(*~
		<docu>
			<summary>
				Provides mechanism for delivering static messages to the supervising applications (SCADA/HMI).	
				<remarks>			
					<note type="important">
						Each messenger has a single placeholder for the message; it stores the most important message from the last context cycle. 
						If there are more messages in a single cycle for the same messenger then less important messages are discarded and replaced by 
						the message with the category of higher severity.							
					</note>
					<note type="important">
						Messenger can send the data to context logger. There is a maximum limit of 10 different messages per messenger in 2 consecutive context cycles.
						The messages that exceed this limit won't be logged when `OnEventRisen` logging is set. 
					    Take this behaviour into account when designing your system.				
					</note>					
				</remarks>			 
			</summary>			
		
		</docu>
~*)
FUNCTION_BLOCK PUBLIC TcoMessenger IMPLEMENTS ITcoMessenger, ITcoMessageProperties, ITcoMessageTextBuilder, ITcoMessageCategorize
VAR			
	(*~
		<docu>
			<summary>
				Most important message of this instance of messenger; stores the most important message from the last context cycle. 
				If there are more messages in a single cycle for the same
				messenger then less important messages are discarded and replaced by the message with the category of higher severity.			 
			</summary>			
		</docu>
	~*)
	_mime : TcoMessage;
	_Parent : ITcoObject;
	{attribute clr [ReadOnly()]}
	_contextIdentity : ULINT;	
	{attribute 'hide'}
	_mds : ARRAY[0..MDS_MAX_INDEX] OF TcoMessageDigest;	
	{attribute 'hide'}
	_condition : eMessageCondition;
	{attribute 'hide'}
	_pinnable : BOOL;		
END_VAR

VAR
	{attribute 'hide'}
	tmpMessageText : STRING(TcoMessengerEnv.MAX_MESSAGE_TEXT_LENGHT);
	{attribute 'hide'}
	refStringBuilder : REFERENCE TO StringBuilder;	
END_VAR

VAR CONSTANT
	MDS_MAX_INDEX : INT := 10;
END_VAR

VAR_STAT
	{attribute 'hide'}
	_conflictingStringBuilder : StringBuilder;
END_VAR

(*~
	<docu>
		<summary>			
			Appends string to the message text. 
		</summary>
		<remarks>
			<note type="warning">
				The size of the resulting string should not be more than '160' characters. The characters exceeding this size will be truncated.
			</note>
		</remarks>
	</docu>	
~*)
{attribute 'hide'}
{attribute 'obsolete' := 'This method must be accessed ITcoMessageTextBuilder interface'} 
METHOD Append : ITcoMessageTextBuilder
VAR_INPUT
	Text : STRING(TcoMessengerEnv.MAX_MESSAGE_TEXT_LENGHT);
END_VAR
THIS^.StringBuilder.Append(Text);
Append := THIS^;
END_METHOD

(*~
	<docu>
		<summary>			
			Appends any value to the message text. 
		</summary>
		<remarks>
			<note type="warning">
				The size of the resulting string should not be more than '160' characters. The characters exceeding this size will be truncated.
			</note>
		</remarks>
	</docu>	
~*)
METHOD AppendAny : ITcoMessageTextBuilder
VAR_INPUT
	Data : ANY;
END_VAR
THIS^.StringBuilder.AppendAny(Data);
AppendAny := THIS^;
END_METHOD

(*~
	<docu>
		<summary>			
			Gets categorization methods for fluent message builder.
		</summary>		
	</docu>	
~*)
{attribute 'hide'}
{attribute 'obsolete' := 'This method must be accessed ITcoMessageTextBuilder interface'} 
METHOD As : ITcoMessageCategorize
As := THIS^;
END_METHOD

(*~
		<docu>
			<summary>
				Categotizes and creates the message as  'debug'.								 
			</summary>		
		</docu>
~*)
{attribute 'hide'}
{attribute 'obsolete' := 'This method must be accessed ITcoMessageCategorize interface'} 
METHOD PUBLIC AsDebug : ITcoMessageProperties
AsDebug := Post(THIS^.StringBuilder.ToString(), eMessageCategory.Debug);
END_METHOD

(*~
		<docu>
			<summary>
				Categotizes and creates the message as  'error'.								 
			</summary>		
		</docu>
~*)

{attribute 'hide'}
{attribute 'obsolete' := 'This method must be accessed ITcoMessageCategorize interface'} 
METHOD PUBLIC AsError : ITcoMessageProperties
AsError := Post(THIS^.StringBuilder.ToString(), eMessageCategory.Error);
END_METHOD

(*~
		<docu>
			<summary>
				Categotizes and creates the message as  'fatal'.								 
			</summary>		
		</docu>
~*)

{attribute 'hide'}
{attribute 'obsolete' := 'This method must be accessed ITcoMessageCategorize interface'} 
METHOD PUBLIC AsFatal : ITcoMessageProperties
AsFatal := Post(THIS^.StringBuilder.ToString(), eMessageCategory.Fatal);
END_METHOD

(*~
		<docu>
			<summary>
				Categotizes and creates the message as  'information'.								 
			</summary>		
		</docu>
~*)

{attribute 'hide'}
{attribute 'obsolete' := 'This method must be accessed ITcoMessageCategorize interface'} 
METHOD PUBLIC AsInfo : ITcoMessageProperties
AsInfo := Post(THIS^.StringBuilder.ToString(), eMessageCategory.Info);
END_METHOD

(*~
		<docu>
			<summary>
				Categotizes and creates the message as  'trace'.								 
			</summary>		
		</docu>
~*)

{attribute 'hide'}
{attribute 'obsolete' := 'This method must be accessed ITcoMessageCategorize interface'} 
METHOD PUBLIC AsTrace : ITcoMessageProperties
AsTrace := Post(THIS^.StringBuilder.ToString(), eMessageCategory.Trace);
END_METHOD

(*~
		<docu>
			<summary>
				Categotizes and creates the message as 'warning'.								 
			</summary>		
		</docu>
~*)

{attribute 'hide'}
{attribute 'obsolete' := 'This method must be accessed ITcoMessageCategorize interface'} 
METHOD PUBLIC AsWarning : ITcoMessageProperties
AsWarning := Post(THIS^.StringBuilder.ToString(), eMessageCategory.Warning);
END_METHOD

(*~
	<docu>
		<summary>			
			Initiates new message text building for this messenger in fluent-like fashion.
		</summary>		
	</docu>	
~*)
METHOD Build : ITcoMessageTextBuilder
THIS^.StringBuilder.Clear();
Build := THIS^;
END_METHOD

(*~
		<docu>
			<summary>
				Adds message of 'catastrophic' category to the message queue.
				Use this category when there is a situation when the device cannot continue operations due to irrecoverable failure.				 
			</summary>		
		</docu>
~*)
METHOD PUBLIC Catastrophic : ITcoMessageProperties
VAR_INPUT
	(*~
		<docu>
			<summary>
				Arbitrary message string.			 
			</summary>			
		</docu>
	~*)
	Message : STRING(TcoMessengerEnv.MAX_MESSAGE_TEXT_LENGHT);
END_VAR
Catastrophic := THIS^.Post(Message, eMessageCategory.Catastrophic);
END_METHOD

(*~
		<docu>
			<summary>
				Clears the message content.
				<remarks>			
					<note type="important">
						This method is exposed for Rpc calls, for testing purposes. Rpc calls of this method must not be used in production code
					</note>
				</remarks>								 
			</summary>		
		</docu>
~*)
{attribute 'TcRpcEnable'}
METHOD Clear
_mime.TimeStamp :=  DT#1970-01-01-00:00;
_mime.Text := '';
_mime.Identity := 0;
_mime.Category := eMessageCategory.All;
_mime.Cycle := 0;	
_mime.PerCycleCount := 0;
_mime.Pinned := FALSE;
END_METHOD

METHOD PROTECTED Compose : TcoMessage
VAR_INPUT
	Text : STRING(TcoMessengerEnv.MAX_MESSAGE_TEXT_LENGHT);
	Category : eMessageCategory;
END_VAR
IF(_Parent <> 0 AND_THEN _Parent.Context <> 0 AND_THEN _Parent.Context.RealTimeClock <> 0) THEN
	Compose.TimeStamp :=  _Parent.Context.RealTimeClock.NowLocal();	
	Compose.Text := Text;
	Compose.Identity := _Parent.Identity;
	Compose.Category := Category;
	Compose.Cycle := _Parent.Context.StartCycleCount;
	Compose.MessageDigest := Digest(Text, THIS^._Parent.Context.Environment.Messaging.MessageDigestMethod);
END_IF;
END_METHOD

(*~
		<docu>
			<summary>
				Adds message of 'critical' category to the message queue.
				Use this category when a critical error occured, that is not recoverable by the means of software (reset/restore) and a detailed inspection is required.				 
			</summary>		
		</docu>
~*)
METHOD PUBLIC Critical : ITcoMessageProperties
VAR_INPUT
	(*~
		<docu>
			<summary>
				Arbitrary message string.			 
			</summary>			
		</docu>
	~*)
	Message : STRING(TcoMessengerEnv.MAX_MESSAGE_TEXT_LENGHT);
END_VAR
Critical := THIS^.Post(Message, eMessageCategory.Critical);
END_METHOD

(*~
		<docu>
			<summary>
				Adds message of 'debug' category to the message queue.	
			    Use when you need to report debug information for you as programmer. 			 
			</summary>		
		</docu>
~*)
METHOD PUBLIC Debug : ITcoMessageProperties
VAR_INPUT
	(*~
		<docu>
			<summary>
				Arbitrary message string.			 
			</summary>			
		</docu>
	~*)
	Message : STRING(TcoMessengerEnv.MAX_MESSAGE_TEXT_LENGHT);
END_VAR
Debug := THIS^.Post(Message, eMessageCategory.Debug);
END_METHOD

METHOD Digest : DWORD
VAR_INPUT
	Text : Tc2_System.T_MaxString;
	inDigestType : eMessageDigestMethod;
END_VAR
CASE inDigestType OF
	eMessageDigestMethod.CRC8 :
		Digest := TcoCRC_8(Text);
	eMessageDigestMethod.CRC16 :
		Digest := TcoCRC_16(Text);
	eMessageDigestMethod.CRC32 :
		Digest := TcoCRC_32(Text);
	ELSE
		Digest := 0;
END_CASE
END_METHOD

(*~
		<docu>
			<summary>
				Adds message of 'error' category to the message queue.
				Use this categoty when there is a failure that cannot be immediately recovered and an intervention is needed. This is typically a situation when a device fails
				to deliver expected result. 
				Do not use this category to report information about failed process like measurement or detection.				 
			</summary>						
		</docu>
~*)
METHOD PUBLIC Error : ITcoMessageProperties
VAR_INPUT
	(*~
		<docu>
			<summary>
				Arbitrary message string.			 
			</summary>			
		</docu>
	~*)
	Message : STRING(TcoMessengerEnv.MAX_MESSAGE_TEXT_LENGHT);
END_VAR
Error := THIS^.Post(Message, eMessageCategory.Error);
END_METHOD

{attribute 'hide'}
METHOD FB_init : BOOL
VAR_INPUT
	bInitRetains : BOOL; // if TRUE, the retain variables are initialized (warm start / cold start)
	bInCopyCode : BOOL;  // if TRUE, the instance afterwards gets moved into the copy code (online change)
	ParentObject : ITcoObject;
END_VAR
_Parent := ParentObject;
_contextIdentity := ParentObject.Identity;
END_METHOD

(*~
		<docu>
			<summary>
				Adds message of 'information' category to the message queue.	
				Use when you want to deliver information to the user, that has only informative character and does not adversely affect a process.			 
			</summary>			
		</docu>
~*)
METHOD PUBLIC Info  : ITcoMessageProperties
VAR_INPUT
	(*~
		<docu>
			<summary>
				Arbitrary message string.			 
			</summary>			
		</docu>
	~*)
	Message : STRING(TcoMessengerEnv.MAX_MESSAGE_TEXT_LENGHT);
END_VAR
Info := THIS^.Post(Message, eMessageCategory.Info);
END_METHOD

METHOD PRIVATE LogMessage 
VAR_IN_OUT
	inMessage : TcoMessage;
END_VAR
VAR
	_index : INT;
	_freeIndex : INT;	
END_VAR
CASE _Parent.Context.Environment.Messaging.MessengerLoggingMethod OF
	eMessengerLogMethod.OnEventRisen :
        IF(_Parent.Context.Environment.Messaging.MessageDigestMethod = eMessageDigestMethod.NONE) THEN
			inMessage.MessageDigest := Digest(inMessage.Text, eMessageDigestMethod.CRC32);
		END_IF
	
		_freeIndex := 0;
		    
		FOR _index := 0 TO MDS_MAX_INDEX DO
			IF(_mds[_index].Cycle = inMessage.Cycle - 1 OR _mds[_index].Cycle = inMessage.Cycle) 
			AND_THEN (_mds[_index].Digest = inMessage.MessageDigest)
			AND_THEN (_mds[_index].Category = inMessage.Category) THEN			
			    _mds[_index].Cycle := inMessage.Cycle;				
				RETURN;											
			END_IF	
			IF((_mds[_index].Cycle <> inMessage.Cycle - 1) 
			   AND (_mds[_index].Cycle <> inMessage.Cycle)) THEN
				_freeIndex := _index;
			END_IF
		END_FOR
		
		IF(_freeIndex <= THIS^.MDS_MAX_INDEX) THEN
			_mds[_freeIndex].Digest := inMessage.MessageDigest;
			_mds[_freeIndex].Cycle := inMessage.Cycle;
			_mds[_freeIndex].Category := inMessage.Category;
			_Parent.Context.Logger.PushMessage(inMessage);		
		END_IF;
	eMessengerLogMethod.Continuous:
	    _Parent.Context.Logger.PushMessage(inMessage);
END_CASE
END_METHOD

(*~
		<docu>
			<summary>
				Adds message of 'notification' category to the message queue.
				Use this category when you want to report a notification that may be of interest to the user, but does not adveresly affect a process.			 
			</summary>				
		</docu>
~*)
METHOD Notify : ITcoMessageProperties
VAR_INPUT
	(*~
		<docu>
			<summary>
				Arbitrary message string.			 
			</summary>			
		</docu>
	~*)
	Message : STRING(TcoMessengerEnv.MAX_MESSAGE_TEXT_LENGHT);
END_VAR
Notify := THIS^.Post(Message, eMessageCategory.Notification);
END_METHOD

METHOD OnCondition : ITcoMessages
VAR_INPUT
	inCondition : BOOL;
END_VAR
IF (inCondition) THEN
	_condition := eMessageCondition.Active;
ELSE
	_condition := eMessageCondition.Inactive;
END_IF

OnCondition := THIS^;
END_METHOD

(*~
	<docu>
		<summary>
			Pins this message that no other message will override it. 
			The messenger won't accept new messages until acknowledged in diagnostics view by user, unipenned by `Unpin()` methods or cleared by `Clear()` method
			of this messenger.						
		</summary>
		<note type="important">
			Pinned messages do no accept incomming messages on the same messenger. The incomming messages will be though the context logger when active.
		</note>
	</docu>
~*)
//~
{attribute 'hide'}
{attribute 'obsolete' := 'This method must be called exclusively over ITcoMessageProperties interface'}
//~ 
METHOD Pin : ITcoMessageProperties
IF(_Parent <> 0 AND_THEN _Parent.Context <> 0) THEN
	IF(_pinnable AND_THEN _mime.Cycle = _Parent.Context.StartCycleCount)THEN
		_mime.Pinned := TRUE;
	END_IF;
END_IF;

Pin := THIS^;
END_METHOD

(*~
	<docu>
		<summary>
			Gets `true` when this messanger is pinned (awaiting acknowledgement in diagnostics view).
		</summary>
	</docu>
~*)
PROPERTY Pinned : BOOL
GET
Pinned := _mime.Pinned AND_THEN tmpMessageText = _mime.Text;
END_GET
END_PROPERTY

(*~
		<docu>
			<summary>
				Creates message of given category for this messenger.				 
			</summary>				
		</docu>
~*)
METHOD PUBLIC Post : ITcoMessageProperties
VAR_INPUT
	(*~
		<docu>
			<summary>
				Arbitrary message string.			 
			</summary>			
		</docu>
	~*)
	Message : STRING(TcoMessengerEnv.MAX_MESSAGE_TEXT_LENGHT);
	(*~
		<docu>
			<summary>
				Message category.			 
			</summary>			
		</docu>
	~*)
	Category : eMessageCategory;	
END_VAR

VAR
	_wouldBeMime : TcoMessage;
END_VAR
Post := THIS^;

tmpMessageText := Message;

_pinnable := FALSE;

IF(_condition = eMessageCondition.Inactive) THEN
	_condition := eMessageCondition.Unconditional;	
	RETURN;
END_IF

_condition := eMessageCondition.Unconditional;


IF(_Parent <> 0 AND_THEN _Parent.Context <> 0 AND_THEN _Parent.Context.Environment <> 0 AND_THEN _Parent.Context.Environment.Messaging <> 0) THEN
	IF(Category < THIS^._Parent.Context.Environment.Messaging.MinLevel
	  OR _Parent.Context.Environment.Messaging.IsSuspended) THEN
		RETURN;
	END_IF; 	
		
	IF (NOT _mime.Pinned) THEN 
		_mime.PerCycleCount := _mime.PerCycleCount + 1;
		_wouldBeMime := Compose(Message, Category);		
		_wouldBeMime.PerCycleCount := _mime.PerCycleCount;		
	ELSIF(_mime.Pinned 
	AND_THEN (_mime.Text <>  Message OR _mime.Category <> Category))
	THEN		
		IF(	_mime.PerCycleCount < 255) THEN	
			_mime.PerCycleCount := _mime.PerCycleCount + 1;	
		END_IF;
	END_IF;		
	
    // Same cycle filter for most important messge.
	IF(_mime.Cycle = _Parent.Context.StartCycleCount) THEN		 	
		IF(_wouldBeMime.Category > _mime.Category) 
		AND (NOT _mime.Pinned) THEN	 
			_mime := _wouldBeMime;
		END_IF;
	ELSE
	// Different cycle					  	    		
		IF (NOT _mime.Pinned) THEN
			_wouldBeMime.PerCycleCount := 1;  													
			_mime := _wouldBeMime;										
		END_IF;
	END_IF;	

	_pinnable := TRUE;
	LogMessage(_wouldBeMime);		
END_IF;
END_METHOD

(*~
		<docu>
			<summary>
				Adds message of 'programming error' category to the message queue.	
				Use this category to inform about a possible programming error, defect in settings or missing information at a level of programming or system or process settings.			 
			</summary>				
		</docu>
~*)
METHOD PUBLIC Programming : ITcoMessageProperties
VAR_INPUT
	(*~
		<docu>
			<summary>
				Arbitrary message string.			 
			</summary>			
		</docu>
	~*)
	Message : STRING(TcoMessengerEnv.MAX_MESSAGE_TEXT_LENGHT);
END_VAR
Programming := THIS^.Post(Message, eMessageCategory.ProgrammingError);
END_METHOD

PROPERTY StringBuilder : REFERENCE TO StringBuilder
GET
VAR
END_VAR

VAR_INST
	_lastCycleAccess : ULINT;
END_VAR
IF(__ISVALIDREF(refStringBuilder)) THEN
	StringBuilder REF= refStringBuilder;
ELSE
	StringBuilder REF= _conflictingStringBuilder;
END_IF
END_GET
END_PROPERTY

(*~
		<docu>
			<summary>
				Adds message of 'trace' category to the message queue.	
				Use when you need to track detailed information about internal states of the program for detailed visibility. 
				This is lowest level of category that can be used in production, for detailed observation of PLC program.			 
			</summary>					
		</docu>
~*)
METHOD PUBLIC Trace : ITcoMessageProperties
VAR_INPUT
	(*~
		<docu>
			<summary>
				Arbitrary message string.			 
			</summary>			
		</docu>
	~*)
	Message : STRING(TcoMessengerEnv.MAX_MESSAGE_TEXT_LENGHT);
END_VAR
Trace := THIS^.Post(Message, eMessageCategory.Trace);
END_METHOD

(*~
	<docu>
		<summary>
			Unpins this messenger.
		</summary>
	</docu>
~*) 
METHOD UnPin
IF (_mime.Pinned) THEN
	IF(_Parent <> 0 AND_THEN _Parent.Context <> 0) THEN
		THIS^.Post('Message unpinned by the controller.', eMessageCategory.Info);
	END_IF;	
END_IF; 
_mime.Pinned := FALSE;
END_METHOD

(*~
		<docu>
			<summary>
				Adds message of 'warning' category to the message queue.
				Use this category when you want to report to the user an information about a possible problem, that may adversly affect a process.
				Information in this cateogory aims to help the user to identify a problem, the cause of such problem does not necessarily stops the process.				 
			</summary>					
		</docu>
~*)
METHOD PUBLIC Warning  : ITcoMessageProperties
VAR_INPUT
	(*~
		<docu>
			<summary>
				Arbitrary message string.			 
			</summary>			
		</docu>
	~*)
	Message : STRING(TcoMessengerEnv.MAX_MESSAGE_TEXT_LENGHT);
END_VAR
Warning := THIS^.Post(Message, eMessageCategory.Warning);
END_METHOD

END_FUNCTION_BLOCK

(* stored: Version 1.1.0.1
   POU TcoMessenger: Id {bb89b26f-ec79-4812-bab7-3579b2b6d1be}, SpecialFunc None
   Folder AsCategory: Id {5e652e11-5ec7-0558-355e-a541dc07128e}
   Folder Messages: Id {56442304-2644-4fe1-b5d1-eb5248dd12e5}
   Folder MessageTextBuilder: Id {84becd26-58f3-0433-37df-29b8ef02e286}
   Method Append: Id {c1ccc337-ea54-00a4-1ba1-6c6567af5ea4}
   Method AppendAny: Id {0a142272-dc83-0b4b-1516-3181619f1e79}
   Method As: Id {4c9973fd-22fb-0755-0689-dcf3cb571511}
   Method AsDebug: Id {9a15fab6-7d2d-0a2a-2268-2662b67885b9}
   Method AsError: Id {ac55723d-e0c1-0cbc-0399-d1c7dedda6ed}
   Method AsFatal: Id {4a4ed82a-2ebf-0f89-3ade-833a0f25d7e7}
   Method AsInfo: Id {4609573e-f820-0eb5-286d-ad5f41802b14}
   Method AsTrace: Id {c619e331-47c0-0a43-09f7-4b71655e3245}
   Method AsWarning: Id {b28d1072-2a77-093a-33e6-3e8a6557022d}
   Method Build: Id {5eccd1dc-e984-03df-06f9-afb4e2349f53}
   Method Catastrophic: Id {3ead99e7-d4fa-03f6-3060-81990c2076df}
   Method Clear: Id {640fefd4-a9aa-0de1-3f5c-cce4bd50449f}
   Method Compose: Id {3447ad14-6768-48d6-b294-87e00174ef1e}
   Method Critical: Id {a9264967-6c30-0c25-362d-a0380aaea992}
   Method Debug: Id {bd0230f7-b5de-4707-ba4a-f8b17cc23976}
   Method Digest: Id {de6a9eab-3c62-0e43-3529-2cc01fda6c4e}
   Method Error: Id {dc14c403-f11e-4200-ac36-567c3d997bf6}
   Method FB_init: Id {23bbd1ba-9be3-4c0b-a177-bc9de93be447}
   Method Info: Id {d1f4840f-86c5-482b-8fb7-443b9b1c585c}
   Method LogMessage: Id {0b6b2fe7-cb26-02a6-0b72-2570a4f5cb53}
   Method Notify: Id {1595dfe7-5719-459e-bdf2-0e7976c85511}
   Method OnCondition: Id {1097de5a-fc1b-0b3c-3c7e-2650c89e121b}
   Method Pin: Id {03e6fdf6-0b38-029d-1385-1c4ef7329d4e}
   Property Pinned: Id {2b9d6a13-0120-0ade-1711-eabdfe133e7e}
   Get Get: Id {922308b3-7383-055d-30c5-1612ea638ab3}
   Method Post: Id {7e1c7e2b-5612-469e-9139-08754fd973ea}
   Method Programming: Id {1f1b6a21-6158-44a7-b79e-b3fcea42c4e1}
   Property StringBuilder: Id {a28ba21a-3e8e-0432-3e41-e8c00eb1332b}
   Get Get: Id {534e9e44-3b1f-00eb-2516-5f0d53690ccd}
   Method Trace: Id {5a17dee2-c171-4127-9ee1-30d4a06a53bf}
   Method UnPin: Id {648f9a53-8d9f-0466-2e58-e936e7aff424}
   Method Warning: Id {dd00674c-7475-44d4-8400-894897951e0b} *)
